PROGRAM MAIN
VAR
END_VAR

// Call I/O Mapping Program
PRG_Mapping();

END_PROGRAM

(* stored: Version 1.1.0.1
   POU MAIN: Id {0ea7724f-a5c0-437c-ab1a-f4a60ea9c49c} *)
